TYPE ST_IsoMon_DeviceSignals :
STRUCT
	insulationResistance_kOhm : REAL;
	minInsulationValue	 	: REAL;
	voltageDCPlusToMinus 	: REAL;
	voltageDCPlusToPE	 	: REAL;
	voltageDCMinusToPE	 	: REAL;
	couplingToSystem	 	: REAL;
	couplingtoEarth		 	: REAL;
	deviceError			 	: REAL;
	deviceInactive			: REAL;
	dcOffset				: REAL;
	measurementQuality		: REAL;
END_STRUCT
END_TYPE

(* stored: Version 1.1.0.1
   DUT ST_IsoMon_DeviceSignals: Id {f7a84d8e-34f8-4a8a-93c5-daa5b778e108} *)
